(* Blister Pack Counter to Target *)

PROGRAM main
  VAR
    FaultEvent AT %IX0.3 : BOOL := 125; (* Various Fault Event Placeholder *)
    Reset AT %IX0.1 : BOOL; (* Internal Reset or External Reset of Counter *)
    MaintenanceAlert AT %QX0.2 : BOOL; (* Detection of Too Many Faults *)
    Force AT %QX0.3 : BOOL; (* Force Reset of Maintenance Alert *)
    Counter : INT; (* Pill Count Variable for SCADA *)
    CTU0 : CTU;
    TOF0 : TOF;
    SR0 : SR;
  END_VAR
  VAR  (* added by the conversion: wires and edge detectors of the diagram *)
    R_TRIG1 : R_TRIG;
  END_VAR

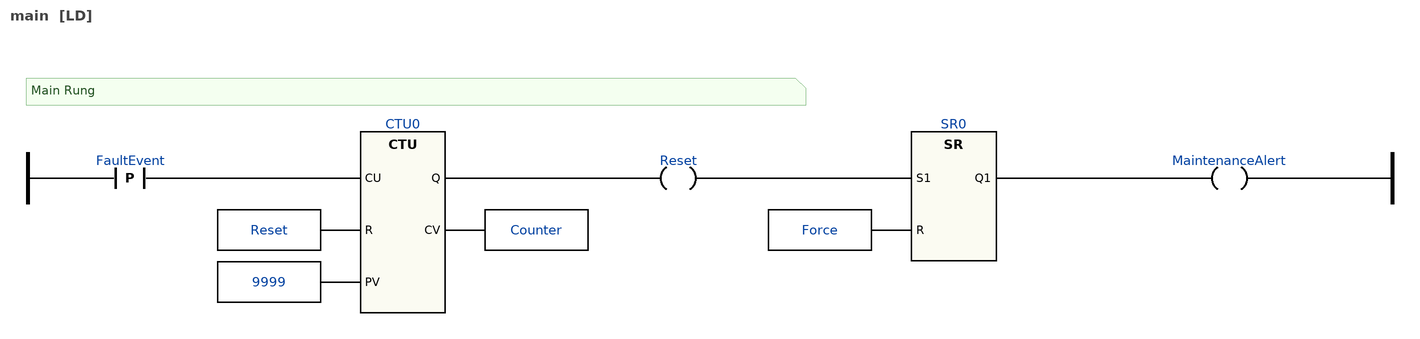
(* LD diagram, written out as Structured Text *)
(* Main Rung *)
R_TRIG1(CLK := FaultEvent);
CTU0(CU := R_TRIG1.Q, R := Reset, PV := 9999);
Reset := CTU0.Q;
SR0(S1 := CTU0.Q, R := Force);
MaintenanceAlert := SR0.Q1;
Counter := CTU0.CV;
END_PROGRAM
